// SIMATIC S7-200 project (STEP 7-Micro/WIN), CPU 226 CN REL 02.01

SYMBOL_TABLE USER1
Sens_Origen      I0.0     // Sensor inductivo de origen para homing del servo
FC_Derecha       I0.1     // Final de carrera derecho limite fisico forward
FC_Izquierda     I0.2     // Final de carrera izquierdo limite fisico reverse
CilV_Abajo       I0.3     // Sensor brazo vertical en posicion abajo
CilV_Arriba      I0.4     // Sensor brazo vertical en posicion arriba
Giro_Izquierda   I0.5     // Sensor actuador rotatorio posicion izquierda antihoraria
Giro_Derecha     I0.6     // Sensor actuador rotatorio posicion derecha horaria
CilDV_Ext        I0.7     // Sensor doble vastago extendido
CilDV_Ret        I1.0     // Sensor doble vastago retraido
Pinza_Cer        I1.1     // Confirmacion de pinza cerrada pieza sujeta
Estado_Servo     I1.2     // Driver servo en estado listo para operar Ready
Btn_Paro         I2.4     // Boton de paro panel de operador
Btn_Marcha       I2.5     // Boton de marcha panel de operador
Seta_Emerg       I2.6     // Seta de emergencia fisica NC
Selector         I2.7     // Selector de modo panel de operador
Servo_Pulsos     Q0.0     // Tren de pulsos PTO para servo motor lineal
Servo_Dir        Q0.2     // Direccion del servo gestionado por MAP_SERV
V_Cil_Vert       Q0.3     // Valvula cilindro vertical brazo arriba
V_Giro_AH        Q0.4     // Valvula actuador rotatorio sentido antihorario
V_Giro_H         Q0.5     // Valvula actuador rotatorio sentido horario
V_Cil_DV         Q0.6     // Valvula doble vastago extendido
V_Pinza_Abre     Q0.7     // Valvula apertura de pinza neumatica
V_Pinza_Cierra   Q1.0     // Valvula cierre de pinza neumatica
Joy_Run_Flag     V29.0    // Bit de marcha de la cinta de transporte
Joy_Dir_Flag     V29.1    // Bit de direccion de la cinta de transporte
Joy_Rot_L_Flag   V29.2    // Bit de giro antihorario del brazo
Joy_Rot_R_Flag   V29.3    // Bit de giro horario del brazo
Joy_Cil_Vert_Flag V29.4    // Bit de cilindro vertical brazo arriba
Joy_Cil_DV_Flag  V29.5    // Bit de cilindro doble vastago extendido
Joy_Grip_Close_Flag V29.6    // Bit de cierre de pinza neumatica
Joy_Grip_Open_Flag V29.7    // Bit de apertura de pinza neumatica
done_modbus      M10.2    // marca done para libreria modbus (init)
error_modbus     VB8      // byte de error para libreria modbus (init)
done_modbus2     M10.3    // marca done para libreria modbus
error_modbus2    VB9      // byte de error para libreria modbus
direccion        V10.1    // direccion de movimiento de la cinta de transporte
error            VB11     // error de la funcion MoveVelocity
c_pos            VD12     // posicion de la funcion MoveVelocity
done_paro        V16.0    // bit de hecho de la funcion Stop
velocidad        VD20     // velocidad para la funcion MoveVelocity
velocidad_buff   VD24     // buffer para la escritura dinamica de la velocidad en MoveVelocity
Servo_C_Pos      VD40     // Posicion actual del servo en pulsos (salida Q0_0_CTRL)
Sol_AP           V0.0     // Solicitud Alimentacion a Procesamiento
Ack_AP           V1.0     // Reconocimiento AP
Sol_PE           V2.0     // Solicitud Procesamiento a Ensamblaje
Ack_PE           V3.0     // Reconocimiento PE
Sol_ES           V4.0     // Solicitud Ensamblaje a Seleccion
Ack_ES           V5.0     // Reconocimiento ES
Ack_MA           V0.1     // Reconocimiento marcha Unidad de Alimentacion
Marcha_A         V1.1     // Solicitud de marcha para la Unidad de Alimentacion
Ack_MP           V2.1     // Reconocimiento marcha Unidad de Procesammiento
Marcha_P         V3.1     // Solicitud de marcha para la Unidad de Procesamiento
Ack_ME           V4.1     // Reconocimiento marcha Unidad de Ensamblaje
Marcha_E         V5.1     // Solicitud de marcha para la Unidad de Ensamblaje
Ack_MS           V6.1     // Reconocimiento marcha Unidad de Seleccion
Marcha_S         V7.1     // Solicitud de marcha para la Unidad de Seleccion
Alim_OK          V0.2     // Unidad de Alimentacion disponible
Proc_OK          V2.2     // Unidad de Procesamiento disponible
Ens_OK           V4.2     // Unidad de Ensamblaje disponible
Sel_OK           V6.2     // Unidad de Seleccion disponible
Pieza_Metal      V6.3     // Pieza identificada por la unidad de seleccion es totalmente metalica
Pieza_Mixta      V6.4     // Pieza identificada por la unidad de seleccion es totalmente mixta
Pieza_Plastica   V6.5     // Pieza identificada por la unidad de seleccion es totalmente plastica
END_SYMBOL_TABLE

SYMBOL_TABLE S7-200 Symbols
Always_On        SM0.0    // 始终接通为 ON
First_Scan_On    SM0.1    // 仅第一个扫描周期中接通为 ON
END_SYMBOL_TABLE

ORGANIZATION_BLOCK MAIN:OB1
TITLE=CONTROL DE VELOCIDAD Y BRAZO CON JOYSTICK - ESTACION DE TRANSPORTE
//  Este programa controla la cinta de transporte y el brazo neumatico manualmente con el joystick.
//  Hace uso de las funciones MoveVelocity (SBR3) y Stop (SBR4) de la libreria MAP_SERV.
BEGIN
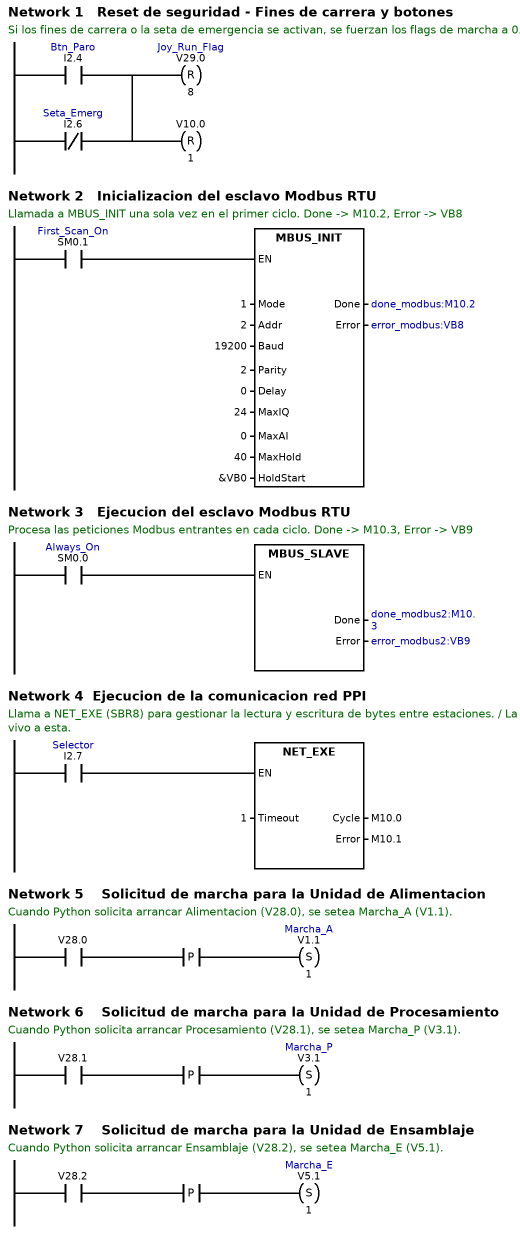
Network 1 //  Reset de seguridad - Fines de carrera y botones
//  Si los fines de carrera o la seta de emergencia se activan, se fuerzan los flags de marcha a 0.
LD     Btn_Paro:I2.4
ON     Seta_Emerg:I2.6
R      Joy_Run_Flag:V29.0, 8
R      V10.0, 1
Network 2 //  Inicializacion del esclavo Modbus RTU
//  Llamada a MBUS_INIT una sola vez en el primer ciclo. Done -> M10.2, Error -> VB8
LD     First_Scan_On:SM0.1
CALL   MBUS_INIT:SBR5, 1, 2, 19200, 2, 0, 24, 0, 40, &VB0, done_modbus:M10.2, error_modbus:VB8
Network 3 //  Ejecucion del esclavo Modbus RTU
//  Procesa las peticiones Modbus entrantes en cada ciclo. Done -> M10.3, Error -> VB9
LD     Always_On:SM0.0
CALL   MBUS_SLAVE:SBR6, done_modbus2:M10.3, error_modbus2:VB9
Network 4 // Ejecucion de la comunicacion red PPI
// Llama a NET_EXE (SBR8) para gestionar la lectura y escritura de bytes entre estaciones.
// La entrada del selector es la que activa esta rutina para poder desactivarla cuando se requiera conectar en vivo a esta.
LD     Selector:I2.7
CALL   NET_EXE:SBR8, 1, M10.0, M10.1
Network 5 //   Solicitud de marcha para la Unidad de Alimentacion
//   Cuando Python solicita arrancar Alimentacion (V28.0), se setea Marcha_A (V1.1).
LD     V28.0
EU
S      Marcha_A:V1.1, 1
Network 6 //   Solicitud de marcha para la Unidad de Procesamiento
//   Cuando Python solicita arrancar Procesamiento (V28.1), se setea Marcha_P (V3.1).
LD     V28.1
EU
S      Marcha_P:V3.1, 1
Network 7 //   Solicitud de marcha para la Unidad de Ensamblaje
//   Cuando Python solicita arrancar Ensamblaje (V28.2), se setea Marcha_E (V5.1).
LD     V28.2
EU
S      Marcha_E:V5.1, 1
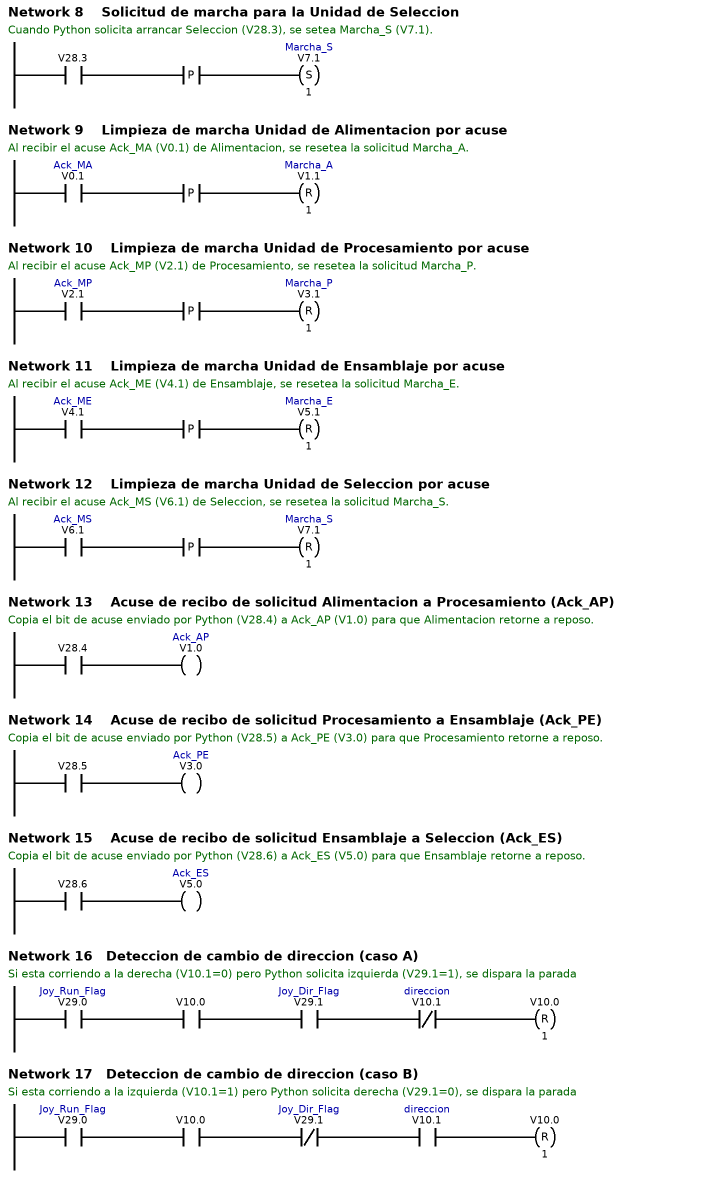
Network 8 //   Solicitud de marcha para la Unidad de Seleccion
//   Cuando Python solicita arrancar Seleccion (V28.3), se setea Marcha_S (V7.1).
LD     V28.3
EU
S      Marcha_S:V7.1, 1
Network 9 //   Limpieza de marcha Unidad de Alimentacion por acuse
//   Al recibir el acuse Ack_MA (V0.1) de Alimentacion, se resetea la solicitud Marcha_A.
LD     Ack_MA:V0.1
EU
R      Marcha_A:V1.1, 1
Network 10 //   Limpieza de marcha Unidad de Procesamiento por acuse
//   Al recibir el acuse Ack_MP (V2.1) de Procesamiento, se resetea la solicitud Marcha_P.
LD     Ack_MP:V2.1
EU
R      Marcha_P:V3.1, 1
Network 11 //   Limpieza de marcha Unidad de Ensamblaje por acuse
//   Al recibir el acuse Ack_ME (V4.1) de Ensamblaje, se resetea la solicitud Marcha_E.
LD     Ack_ME:V4.1
EU
R      Marcha_E:V5.1, 1
Network 12 //   Limpieza de marcha Unidad de Seleccion por acuse
//   Al recibir el acuse Ack_MS (V6.1) de Seleccion, se resetea la solicitud Marcha_S.
LD     Ack_MS:V6.1
EU
R      Marcha_S:V7.1, 1
Network 13 //   Acuse de recibo de solicitud Alimentacion a Procesamiento (Ack_AP)
//   Copia el bit de acuse enviado por Python (V28.4) a Ack_AP (V1.0) para que Alimentacion retorne a reposo.
LD     V28.4
=      Ack_AP:V1.0
Network 14 //   Acuse de recibo de solicitud Procesamiento a Ensamblaje (Ack_PE)
//   Copia el bit de acuse enviado por Python (V28.5) a Ack_PE (V3.0) para que Procesamiento retorne a reposo.
LD     V28.5
=      Ack_PE:V3.0
Network 15 //   Acuse de recibo de solicitud Ensamblaje a Seleccion (Ack_ES)
//   Copia el bit de acuse enviado por Python (V28.6) a Ack_ES (V5.0) para que Ensamblaje retorne a reposo.
LD     V28.6
=      Ack_ES:V5.0
Network 16 //  Deteccion de cambio de direccion (caso A)
//  Si esta corriendo a la derecha (V10.1=0) pero Python solicita izquierda (V29.1=1), se dispara la parada
LD     Joy_Run_Flag:V29.0
A      V10.0
A      Joy_Dir_Flag:V29.1
AN     direccion:V10.1
R      V10.0, 1
Network 17 //  Deteccion de cambio de direccion (caso B)
//  Si esta corriendo a la izquierda (V10.1=1) pero Python solicita derecha (V29.1=0), se dispara la parada
LD     Joy_Run_Flag:V29.0
A      V10.0
AN     Joy_Dir_Flag:V29.1
A      direccion:V10.1
R      V10.0, 1
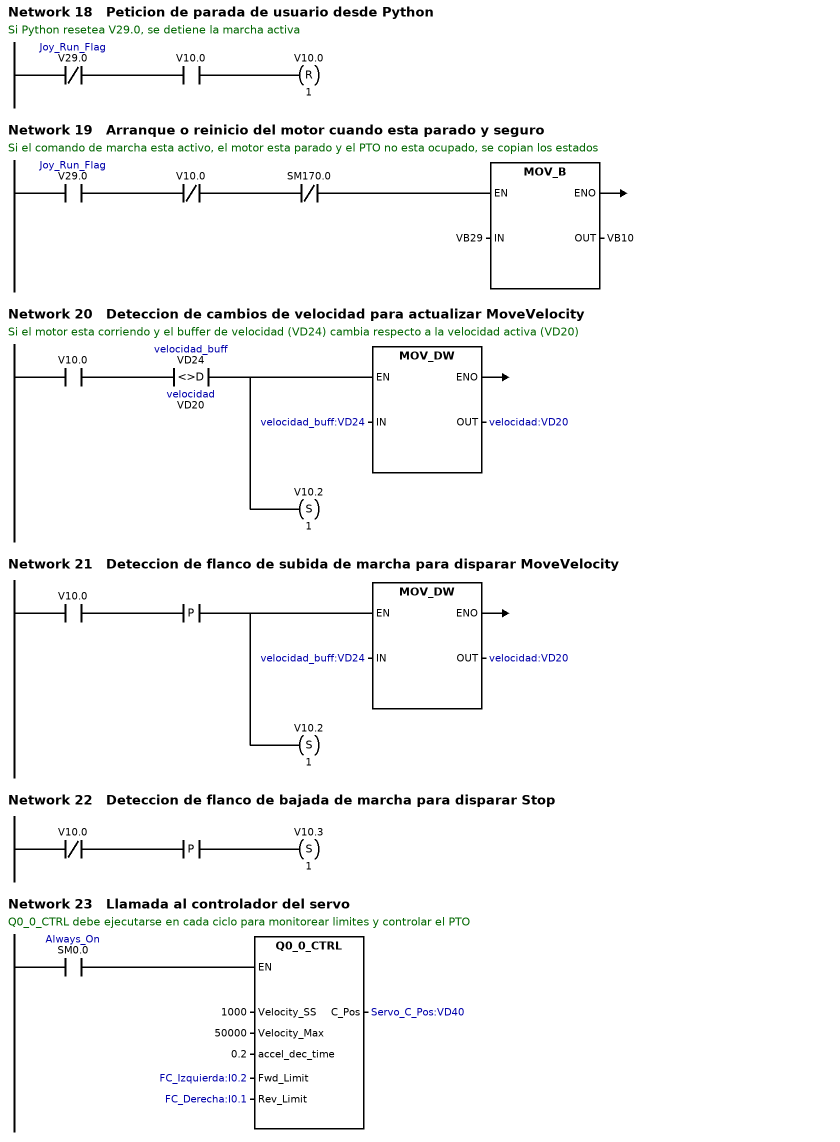
Network 18 //  Peticion de parada de usuario desde Python
//  Si Python resetea V29.0, se detiene la marcha activa
LDN    Joy_Run_Flag:V29.0
A      V10.0
R      V10.0, 1
Network 19 //  Arranque o reinicio del motor cuando esta parado y seguro
//  Si el comando de marcha esta activo, el motor esta parado y el PTO no esta ocupado, se copian los estados
LD     Joy_Run_Flag:V29.0
AN     V10.0
AN     SM170.0
MOVB   VB29, VB10
Network 20 //  Deteccion de cambios de velocidad para actualizar MoveVelocity
//  Si el motor esta corriendo y el buffer de velocidad (VD24) cambia respecto a la velocidad activa (VD20)
// Solicita pulso de ejecucion de MoveVelocity
LD     V10.0
AD<>   velocidad_buff:VD24, velocidad:VD20
MOVD   velocidad_buff:VD24, velocidad:VD20
S      V10.2, 1
Network 21 //  Deteccion de flanco de subida de marcha para disparar MoveVelocity
// Solicita pulso de ejecucion de MoveVelocity
LD     V10.0
EU
MOVD   velocidad_buff:VD24, velocidad:VD20
S      V10.2, 1
Network 22 //  Deteccion de flanco de bajada de marcha para disparar Stop
// Solicita pulso de ejecucion de Stop
LDN    V10.0
EU
S      V10.3, 1
Network 23 //  Llamada al controlador del servo
//  Q0_0_CTRL debe ejecutarse en cada ciclo para monitorear limites y controlar el PTO
LD     Always_On:SM0.0
CALL   Q0_0_CTRL:SBR1, 1000, 50000, 0.2, FC_Izquierda:I0.2, FC_Derecha:I0.1, Servo_C_Pos:VD40
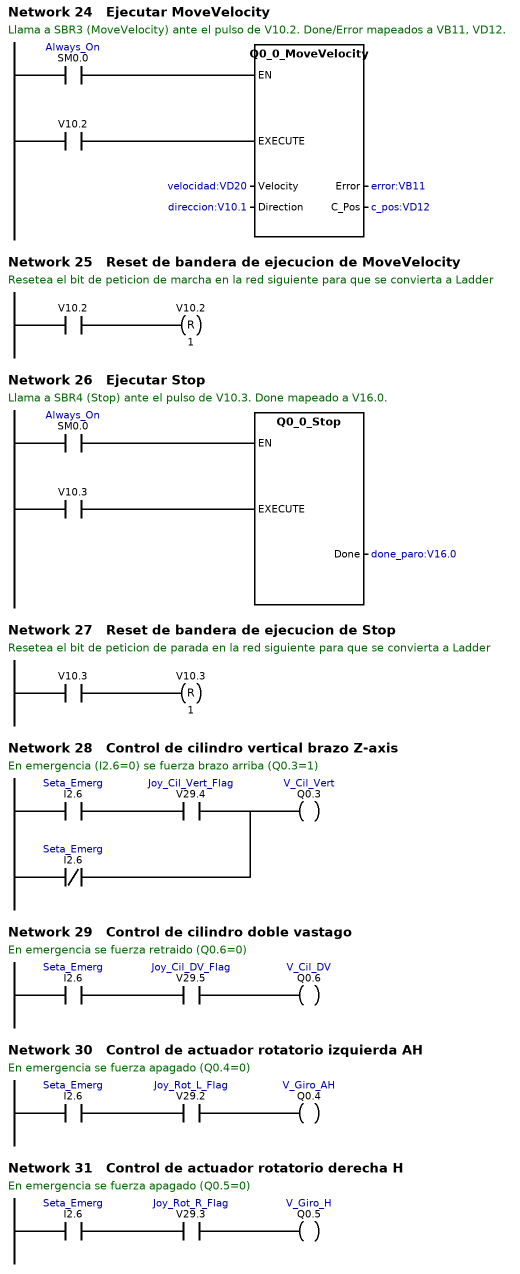
Network 24 //  Ejecutar MoveVelocity
//  Llama a SBR3 (MoveVelocity) ante el pulso de V10.2. Done/Error mapeados a VB11, VD12.
LD     Always_On:SM0.0
=      L60.0
LD     V10.2
=      L63.7
LD     L60.0
CALL   Q0_0_MoveVelocity:SBR3, L63.7, velocidad:VD20, direccion:V10.1, error:VB11, c_pos:VD12
Network 25 //  Reset de bandera de ejecucion de MoveVelocity
//  Resetea el bit de peticion de marcha en la red siguiente para que se convierta a Ladder
LD     V10.2
R      V10.2, 1
Network 26 //  Ejecutar Stop
//  Llama a SBR4 (Stop) ante el pulso de V10.3. Done mapeado a V16.0.
LD     Always_On:SM0.0
=      L60.0
LD     V10.3
=      L63.7
LD     L60.0
CALL   Q0_0_Stop:SBR4, L63.7, done_paro:V16.0
Network 27 //  Reset de bandera de ejecucion de Stop
//  Resetea el bit de peticion de parada en la red siguiente para que se convierta a Ladder
LD     V10.3
R      V10.3, 1
Network 28 //  Control de cilindro vertical brazo Z-axis
//  En emergencia (I2.6=0) se fuerza brazo arriba (Q0.3=1)
LD     Seta_Emerg:I2.6
A      Joy_Cil_Vert_Flag:V29.4
ON     Seta_Emerg:I2.6
=      V_Cil_Vert:Q0.3
Network 29 //  Control de cilindro doble vastago
//  En emergencia se fuerza retraido (Q0.6=0)
LD     Seta_Emerg:I2.6
A      Joy_Cil_DV_Flag:V29.5
=      V_Cil_DV:Q0.6
Network 30 //  Control de actuador rotatorio izquierda AH
//  En emergencia se fuerza apagado (Q0.4=0)
LD     Seta_Emerg:I2.6
A      Joy_Rot_L_Flag:V29.2
=      V_Giro_AH:Q0.4
Network 31 //  Control de actuador rotatorio derecha H
//  En emergencia se fuerza apagado (Q0.5=0)
LD     Seta_Emerg:I2.6
A      Joy_Rot_R_Flag:V29.3
=      V_Giro_H:Q0.5
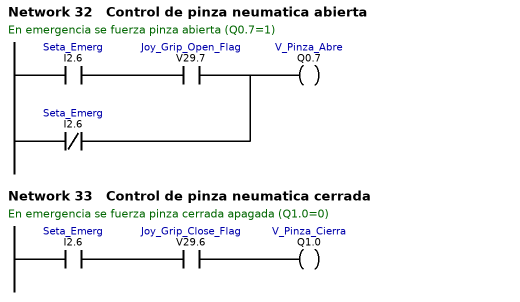
Network 32 //  Control de pinza neumatica abierta
//  En emergencia se fuerza pinza abierta (Q0.7=1)
LD     Seta_Emerg:I2.6
A      Joy_Grip_Open_Flag:V29.7
ON     Seta_Emerg:I2.6
=      V_Pinza_Abre:Q0.7
Network 33 //  Control de pinza neumatica cerrada
//  En emergencia se fuerza pinza cerrada apagada (Q1.0=0)
LD     Seta_Emerg:I2.6
A      Joy_Grip_Close_Flag:V29.6
=      V_Pinza_Cierra:Q1.0
END_ORGANIZATION_BLOCK

// SBR1: protected block, not included

// SBR2: protected block, not included

// SBR3: protected block, not included

// SBR4: protected block, not included

// SBR5: protected block, not included

// SBR6: protected block, not included

// SBR7: protected block, not included

// SBR8: protected block, not included
